Yaskawa INFORM job: EDGEPRO.JBI

/JOB
//NAME EDGEPRO
//POS
///NPOS 3,0,3,0,0,0
///TOOL 9
///POSTYPE PULSE
///PULSE
C00000=0,0,0
C00001=0,0,0
C00002=0,0,0
EC00000=0
EC00001=0
EC00002=0
//INST
<volatile>
///COMM Generated using RoboDK
///ATTR SC,RW
///GROUP1 RB1
NOP
'Program generated by RoboDK v
'6.0.7 for Yaskawa Motoman EPL
'160 on XX/XX/XXXX 18:00:00
'Using nominal kinematics.
'Using Frame Edge (targets wrt
' base):
'100.5,-200.2,300.1,30.0,-20.0
',10.0
'Tool Tool Edge should be clos
'e to:
'-1.5,2.2,99.9,180.0,45.0,-90.
'0
MOVJ C00000 VJ=33.33  +MOVJ EC00000 VJ=100.00
MOVL C00001 V=123.5 PL=8  +MOVJ EC00001 VJ=100.00
PAUSE
TIMER T=1.23
MSG "A long message with "quot"
MSG "es", 'apostrophes' & symb"
MSG "ols: <>[]{}()=+-*/%;#@! a"
MSG "nd more text to make it l"
MSG "onger than eighty charact"
MSG "ers"
'Comment with ; semicolon
DOUT Gripper ON
DOUT OT#(12) OFF
DOUT Pressure ON
WAIT PartPresent=ON T=0.25
WAIT IN#(7)=1
CALL JOB:DOSOMET
x = 1
MOVJ C00002 VJ=33.33 PL=8  +MOVJ EC00002 VJ=100.00
END
